TYPE "ST_TimingRow"
VERSION : 0.1
   STRUCT
      "Id" : DInt;
      "Label" : String[120];
      "TimeClass" : DInt;
      "Count" : UDInt;
      "Last" : Time;
      "Minimum" : Time;
      "Maximum" : Time;
      "Avg" : Time;
   END_STRUCT;
END_TYPE
